{attribute 'qualified_only'}
{attribute 'strict'}
TYPE E_TurCtl : 
(
	e_1 := 1, (*ROSCO*)
	e_2 := 2 (*Lio*)
) SINT;
END_TYPE

(* stored: Version 1.1.0.1
   DUT E_TurCtl: Id {443a4033-2749-42cb-b5fb-22284c015218} *)
